(* IEC 61131-3 sources: PLC_Gen_Frame/Agents4PLC_release/results/task_1778471347, 1 file *)

(* ---- output.ST ---- *)
FUNCTION_BLOCK in
VAR_INPUT
    SoilMoistureSensor1 : REAL;
    SoilMoistureSensor2 : REAL;
    WeatherForecast : INT;
END_VAR
VAR_OUTPUT
    WaterPump : BOOL;
END_VAR

// Generated by DummyPLCGenerator

END_FUNCTION_BLOCK
